FUNCTION_BLOCK ParamLabelAtLeftEdge (* Parameter value labels at the left edge and an instance name wider than its block at the right edge of a network wider than the minimum network width *)
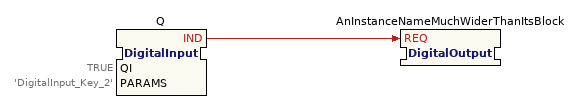
  FBS
    Q : DigitalInput(QI := TRUE, PARAMS := 'DigitalInput_Key_2');
    AnInstanceNameMuchWiderThanItsBlock : DigitalOutput;
  END_FBS
  EVENT_CONNECTIONS
    Q.IND TO AnInstanceNameMuchWiderThanItsBlock.REQ;
  END_CONNECTIONS
END_FUNCTION_BLOCK
